(* IEC 61131-3 sources: LASAL/Class/SafetyCDIAS_Base (part 3) *)

	end_if;

END_FUNCTION

FUNCTION VIRTUAL SafetyCDIAS_Base::GetModuleID
	VAR_OUTPUT
		ud_ModuleID 	: UDINT;
	END_VAR

  // no module
  ud_ModuleID := 16#ff;

END_FUNCTION

FUNCTION VIRTUAL GLOBAL SafetyCDIAS_Base::Init
  VAR
		MyPara 	  : CmdStruct;
		MyResult	: results;
  END_VAR

//============================ Profiler start======================================================
#ifdef DM_Profiler
  InitTimeMeasurement(usMode := DMTIME_RT);
  InitTimeMeasurement(usMode := DMTIME_CY);
  InitTimeMeasurement(usMode := DMTIME_RTPOSTSCAN);
#endif
//============================ Profiler end========================================================

#ifdef DEACTIVATED_LSL
  IF Place.Read() = DEACTIVATED_LSL THEN
    State.uiIO_Flags                  := 0;
    State.uiIO_Flags.NoHW             := 1;
    State.uiIO_Flags.PhysicAccessOff  := 1;
    return;
  END_IF;
#endif

  case InitStep of
    0:
      // initialize HwBaseCDIAS
      if InitSafetyBase() then
        InitStep += 1;
      else
        //Remember flag that init failed, we must not try again otherwise the local var pSafetyManagerThis gets overwritten with nil if it already has been initialized
        InitStep := -1;
      end_if;

    1:
      // add update tasks in dependence on priority (prio 1 is added when us_FirstScan = 2, prio 2 @ us_FirstScan = 3...)
      if ( ( us_FirstScan - 1 ) = GetTaskPriority() ) then

        AddSafetyTask();

        InitStep += 1;

      end_if;

   2:
      // initialize safety module specific data (cpu, input, output) in last init and send OK to CPU

      if ((us_FirstScan = 10) & ((State.uiIO_Flags = 0 | DelayedStartup = 1))) then

        // log in to safety manager, if there is one
        if pSafetyManagerThis then
          MyPara.uiCmd    := CMD_SM_ADD_MODULE;
          MyPara.aPara[0] := ud_MyModuleID$DINT;
          MyPara.aPara[1] := THIS$DINT;
          pSafetyManagerThis^.NewInst(#MyPara, #MyResult);

          // check if quit error is avaialble
          MyPara.uiCmd    := CMD_SM_QUIT_ERROR_AVAILABLE;
          MyPara.aPara[0] := THIS$DINT;
          pSafetyManagerThis^.NewInst(#MyPara, #MyResult);

          // if the DLL has been found and the version shows that CDIAS safety is supported
          b_QuitErrorAvailable := (MyResult.aData[0]$DINT <> 0) & (MyResult.aData[4]$UDINT >= SAFETY_DLL_VERSION_CDIAS_QE);

          // give the manager more details about the module (if it didn't work at the first time and the safety number is valid)
          if (b_SafetyInfoOK = FALSE & ((DelayedStartup = 0) | ((DelayedStartup = 1 & SafetyNumber)))) then

            MyPara.uiCmd    := CMD_SM_ADD_MODULE_INFO;
            MyPara.aPara[0] := THIS$DINT;
            MyPara.aPara[1] := SafetyNumber$DINT;
            MyPara.aPara[2] := FW_Version$DINT;
            MyPara.aPara[3] := FPGA_Version$DINT;
            MyPara.aPara[4] := to_DINT(p_ObjectPath^$USINT) + 1; // size of path (length + 1 for the length information)
            MyPara.aPara[5] := p_ObjectPath$DINT;
            pSafetyManagerThis^.NewInst(#MyPara, #MyResult);
            b_SafetyInfoOK := MyResult.aData[0];
          end_if;
        else
          // if there is no manager, we don't have to wait in cywork until the initialisation is finished
          b_ManagerInitialisationFinished := TRUE;
          b_ManagerReadyForSDO            := TRUE;
        end_if;

        InitSafeModule();
      end_if;

    -1:
      //Error, nothing to do here, states are set before

  end_case;

  us_FirstScan += 1;

END_FUNCTION

FUNCTION VIRTUAL SafetyCDIAS_Base::GetTaskPriority
	VAR_OUTPUT
		us_TaskPriority 	: USINT;
	END_VAR

  // highest = default-priority (no change in update order)
  us_TaskPriority := 0;

END_FUNCTION

FUNCTION VIRTUAL SafetyCDIAS_Base::InitSafeModule
	VAR_OUTPUT
		sd_retval 	: DINT;
	END_VAR

  sd_retval := 0;

END_FUNCTION

FUNCTION VIRTUAL SafetyCDIAS_Base::StartDO
  VAR
  	i : DINT;
  END_VAR

  if b_PayloadSupport = FALSE then
    //set right address of do
    MasterConnect.SetNewDOAddressRd( p_data := pPDOReadData$^DINT, ud_address:= ( ui_MyPlace + OFFSET_SPDO_DATA ) );
  end_if;

  //start data object
  MasterConnect.ResetDO( p_data_object := p_HandlePDORead$^DINT, us_state := VARAN_DO_NO_RUN, ud_bytes := MaxLengthPDORead );

  // only for modules with outputs
  if Kennung <> CSDI16x_ID then
    if b_PayloadSupport = FALSE then
      //set right address of do
      MasterConnect.SetNewDOAddressWr( p_data := pPDOWriteData$^DINT, ud_address:= ( ui_MyPlace + OFFSET_SPDO_DATA ) );
    end_if;
    //start data object
    MasterConnect.ResetDO( p_data_object := p_HandlePDOWrite$^DINT, us_state := VARAN_DO_NO_RUN, ud_bytes := MaxLengthPDOWrite);

    if (AdditionalSPDOs > 0) then
      for i := 0 to (AdditionalSPDOs-1) do
        if b_PayloadSupport = FALSE then
          //set right address of do
          MasterConnect.SetNewDOAddressWr( p_data := aAdditionalPDOs[i].pPDOWriteData$^DINT, ud_address:= ( ui_MyPlace + OFFSET_SPDO_DATA ) );
        end_if;
        //start data object
        MasterConnect.ResetDO( p_data_object := aAdditionalPDOs[i].p_HandlePDOWrite$^DINT, us_state := VARAN_DO_NO_RUN, ud_bytes := MaxLengthPDOWrite);
      end_for;
    end_if;
  end_if;

  if b_PayloadSupport = FALSE then
    //set right address of do
    MasterConnect.SetNewDOAddressRd(p_data := p_us_Handle_TDO_Read$^DINT, ud_address := ui_MyPlace + OFFSET_STDO_DATA);

    //set right address of do
    MasterConnect.SetNewDOAddressWr(p_data := p_us_Handle_TDO_Write$^DINT, ud_address := ui_MyPlace + OFFSET_STDO_DATA);

    //set right address of do
    MasterConnect.SetNewDOAddressRd(p_data := p_ud_Handle_LED$^DINT, ud_address := ui_MyPlace + OFFSET_LED );
  end_if;

	//start data object
  MasterConnect.ResetDO( p_data_object := p_HandleTDORead$^DINT, us_state := VARAN_DO_NO_RUN, ud_bytes := STDO_LENGTH );

  //start data object
  MasterConnect.ResetDO( p_data_object := p_HandleTDOWrite$^DINT, us_state := VARAN_DO_NO_RUN, ud_bytes := STDO_LENGTH );

	//start data object
	MasterConnect.ResetDO( p_data_object := p_HandleLED$^DINT, us_state := VARAN_DO_CONT_RUN, ud_bytes := 15 );

  // only for modules with outputs
  if Kennung <> CSDI16x_ID then
    if b_PayloadSupport = FALSE then
      //set right address of do
      MasterConnect.SetNewDOAddressWr(p_data := p_ui_UnsafeOutWrite$^DINT, ud_address := ui_MyPlace + OFFSET_UNSAFE_VAR);
    end_if;
    //start data object
    MasterConnect.ResetDO( p_data_object := p_HandleUnsafeOutWrite$^DINT, us_state := VARAN_DO_NO_RUN, ud_bytes := UNSAFE_OUT_LENGTH );
  end_if;

  // fast unsafe variables (only if activated)
  if ActivateFastUnsafeIOs then
    if b_PayloadSupport = FALSE then
      //set right address of do
      MasterConnect.SetNewDOAddressRdWr(p_data:=p_us_Handle_FastUnsafeInputs$^DINT, ud_address_read:=ui_MyPlace + OFFSET_FAST_UNSAFE_IOS, ud_address_write:=ui_MyPlace + OFFSET_FAST_UNSAFE_IOS);
    end_if;
    //start data object
    MasterConnect.ResetDO( p_data_object := p_HandleFastUnsafeIOs$^DINT, us_state := VARAN_DO_CONT_RUN, ud_bytes := 1 );
  end_if;

  if b_PayloadSupport = FALSE then
    //set right address of do
    MasterConnect.SetNewDOAddressWr(p_data := p_us_Handle_TimeSyncHS_Write$^DINT, ud_address := ui_MyPlace + OFFSET_TIMESYNC_HANDSHAKE);
  end_if;
  //start data object
  MasterConnect.ResetDO( p_data_object := p_Handle_TimeSyncHS_Write$^DINT, us_state := VARAN_DO_NO_RUN, ud_bytes := 1 );

END_FUNCTION

FUNCTION VIRTUAL SafetyCDIAS_Base::StopDO
  VAR
  	i : DINT;
  END_VAR

  // stop data objects
	MasterConnect.ResetDO( p_data_object := p_HandlePDORead$^DINT, us_state := VARAN_DO_NO_RUN, ud_bytes := MaxLengthPDORead);

  // only for modules with outputs
  if Kennung <> CSDI16x_ID then

    MasterConnect.ResetDO( p_data_object := p_HandlePDOWrite$^DINT, us_state := VARAN_DO_NO_RUN, ud_bytes := MaxLengthPDOWrite);

    if (AdditionalSPDOs > 0) then
      for i := 0 to (AdditionalSPDOs-1) do
        if b_PayloadSupport = FALSE then
          //set right address of do
          MasterConnect.SetNewDOAddressWr( p_data := aAdditionalPDOs[i].pPDOWriteData$^DINT, ud_address:= ( ui_MyPlace + OFFSET_SPDO_DATA ) );
        end_if;
        //start data object
        MasterConnect.ResetDO( p_data_object := aAdditionalPDOs[i].p_HandlePDOWrite$^DINT, us_state := VARAN_DO_NO_RUN, ud_bytes := MaxLengthPDOWrite);
      end_for;
    end_if;
  end_if;

	MasterConnect.ResetDO( p_data_object := p_HandleTDORead$^DINT, us_state := VARAN_DO_NO_RUN, ud_bytes := STDO_LENGTH );
  b_DOIsRunningTDORead          := 0;

	MasterConnect.ResetDO( p_data_object := p_HandleTDOWrite$^DINT, us_state := VARAN_DO_NO_RUN, ud_bytes := STDO_LENGTH );
  b_DOIsRunningTDOWrite         := 0;

  MasterConnect.ResetDO( p_data_object := p_HandleLED$^DINT, us_state := VARAN_DO_NO_RUN, ud_bytes := 15 );

  MasterConnect.ResetDO( p_data_object := p_Handle_TimeSyncHS_Write$^DINT, us_state := VARAN_DO_NO_RUN, ud_bytes := 1 );
  b_DOIsRunning_TimeSyncHS      := 0;

  // only for modules with outputs
  if Kennung <> CSDI16x_ID then
    MasterConnect.ResetDO( p_data_object := p_HandleUnsafeOutWrite$^DINT, us_state := VARAN_DO_NO_RUN, ud_bytes := UNSAFE_OUT_LENGTH );
    b_DOIsRunningUnsafeOutWrite := 0;
  end_if;

END_FUNCTION

FUNCTION VIRTUAL SafetyCDIAS_Base::InitBuffers
	VAR_OUTPUT
		sd_retval 	: DINT;
	END_VAR

  sd_retval := -1;

  //allocate memory for outgoing SDO (one SDO possible)
  p_SDOOutputBuffer$^void := To_StdLib.Malloc(size := SDO_MAX_LENGTH);

  if ( p_SDOOutputBuffer = NIL ) then
    State.uiIO_Flags				          := 0;
		State.uiIO_Flags.PhysicAccessOff  := 1;
    ClassState := _MemAllocFailed;
    return;
  end_if;

  //allocate memory for incoming SDO list (number of SDO is dynamical)
  //following elements will be added dynamical

  //allocate list
  InputBufferAllocatedNo := SDO_BUFFER_ALLOC_BLOCK;
  p_SDOInputBuffer$^void := To_StdLib.Malloc(size := InputBufferAllocatedNo * SDO_MAX_LENGTH);

  if ( p_SDOInputBuffer = NIL ) then
    State.uiIO_Flags				          := 0;
		State.uiIO_Flags.PhysicAccessOff  := 1;
    ClassState := _MemAllocFailed;
    return;
  end_if;

  //all buffers initialized
  sd_retval := 0;

END_FUNCTION

FUNCTION VIRTUAL SafetyCDIAS_Base::GetSafetyNumber
	VAR_OUTPUT
		sd_retval 	: DINT;
	END_VAR
  VAR
  	TempPathInfo: PathInfoType;
		MyPara 	    : CmdStruct;
		MyResult	  : results;
  END_VAR

  sd_retval := SDOStdRequ ( us_Command      := SDO_COMMAND_GET_SAFENBR
                          , p_us_RespData   := ( #SafetyNumber )$^USINT
                          , us_RespLength   := sizeof(SafetyNumber)
                          );

  if ( sd_retval <> 0 ) then
    State.uiIO_Flags				          := 0;
		State.uiIO_Flags.PhysicAccessOff  := 1;

    LogError("@ZZZZ (SafetyCDIAS_Base::GetSafetyNumber) No Safety Number available!");
  elsif pConfigMem then
    // store safety number in config memory
    pConfigMem^$HDINT := SafetyNumber;
  end_if;

  sd_retval := SDOStdRequ ( us_Command      := SDO_COMMAND_GET_FW_VERSION
                          , p_us_RespData   := ( #FirmwareVersion )$^USINT
                          , us_RespLength   := sizeof(FirmwareVersionType)
                          );

  if ( sd_retval = 0 ) then
    FW_Version := FirmwareVersion.RevMinor OR (FirmwareVersion.RevMajor SHL 16);

    // Minor Versions starting with 9xxx mark Bootloader versions
    if (FirmwareVersion.RevMinor >= 9000) & (FirmwareVersion.RevMinor < 10000) then
      LogError("@ZZZZ (SafetyCDIAS_Base::GetSafetyNumber) Bootloader version of safety firmware detected! Download a firmware or contact Sigmatek Support!");
    end_if;

    // if we are connected over mover maybe the second try to read the fw version succeeds after the first failed
    if (sd_VaranType = 2) & (ClassState = _ReadFWVerFailed) then
      ClassState := _WaitForSynchronicity;
    end_if;
  else
    State.uiIO_Flags				          := 0;
    State.uiIO_Flags.PhysicAccessOff  := 1;
    ClassState := _ReadFWVerFailed;
    LogError("@ZZZZ (SafetyCDIAS_Base::GetSafetyNumber) No Firmware Version available!");
  end_if;

  InitPathInfo(#TempPathInfo);

  // add own safety number to routing table
  sd_retval := AddRoutingElement( ud_SafeNumber       := SafetyNumber
                                , ud_thisp            := this$UDINT
                                , pObject             := #TempPathInfo
                                );

  // give the manager more details about the module
  if pSafetyManagerThis then
    if ((SafetyNumber & DelayedStartup = 1) | DelayedStartup = 0) then
      MyPara.uiCmd    := CMD_SM_ADD_MODULE_INFO;
      MyPara.aPara[0] := THIS$DINT;
      MyPara.aPara[1] := SafetyNumber$DINT;
      MyPara.aPara[2] := FW_Version$DINT;
      MyPara.aPara[3] := FPGA_Version$DINT;
      MyPara.aPara[4] := to_DINT(p_ObjectPath^$USINT) + 1; // size of path (length + 1 for the length information)
      MyPara.aPara[5] := p_ObjectPath$DINT;
      pSafetyManagerThis^.NewInst(#MyPara, #MyResult);
      b_SafetyInfoOK := MyResult.aData[0];
    end_if;
  else
    // if there is no safety manager, it can only work if old modules are being used (new need the time sync token)

    // if the FPGA Version is lower than 1.4 or the minor firmware version is lower than 100 everything is fine
    if (FPGA_Version < 16#14) | (FW_Version$UINT < 100) then
      // new classes with old modules and without safety manager (hwcontrol) => no problem
    else
      // new classes with new modules and without safety manager (hwcontrol) => problem: noone there to pass on the time sync token
      LogError("@ZZZZ (SafetyCDIAS_Base::GetSafetyNumber) For new safety modules an object of HwControl is needed for time synchronisation!");
    end_if;
  end_if;

END_FUNCTION

FUNCTION SafetyCDIAS_Base::SafetyCDIAS_Base
	VAR_OUTPUT
		ret_code 	: ConfStates;
	END_VAR

#ifdef HWC_LogInit
  HWC_LogInit();
#endif

  //get interface for safety functions
  if ( OS_CILGET(INTERFACE_SAFETY, #pISafety)) then
    pISafety := NIL;

    LogError("@ZZZZ (SafetyCDIAS_Base::SafetyCDIAS_Base) No Safety Interface found!");

  end_if;

  // initialize it with FALSE, if there is anything on local CDIAS it will change to TRUE
  b_SafetyOnLocalCDIAS := FALSE;

  // initialize module count with 0
  ModuleSyncNo := 0;

  ret_code := C_OK;

END_FUNCTION

FUNCTION VIRTUAL GLOBAL SafetyCDIAS_Base::UpDateRT
	VAR_INPUT
		Handle 	      : UDINT;
	END_VAR
  VAR
    PDOLength     : USINT;
    p_ReceiveObj  : pVirtualBase;
    p_addressRd   : ^VaranDOSettingsRd;
    i             : DINT;
		MyPara 	      : CmdStruct;
		MyResult	    : results;
    bValidTDO     : BOOL;
  END_VAR

//============================ Profiler start======================================================
#ifdef  DM_Profiler
  StartTimeMeasurement(usMode := DMTIME_RT);
#endif
//============================ Profiler end========================================================

  // do tdo/pdo communication only, if module has been found and initialized correctly and if there are some LEDs on (else a FW-Update is running)
  if ( State.uiIO_Flags = 0 ) &
     (( ClassState = _SafetyClassOK ) | ( ClassState = _WaitForSynchronicity ) | ( ClassState = _ReinitConfig ) | ( ClassState = _ModFromCfgNotFound ) | ( ClassState = _UnknownCfgError ) | ( ClassState = _UnsafeVarNotFound )) then

    if StartRtDOs then
      if StartRtDOs = 2 then
        //start DOs
        StartDO();
      else
        if b_PayloadSupport = FALSE then
          //set right address of do
          MasterConnect.SetNewDOAddressRd( p_data := pPDOReadData$^DINT, ud_address:= ( ui_MyPlace + OFFSET_SPDO_DATA ) );
        end_if;

        //start data object
        MasterConnect.ResetDO( p_data_object := p_HandlePDORead$^DINT, us_state := VARAN_DO_NO_RUN, ud_bytes := MaxLengthPDORead );
      end_if;

      StartRtDOs := 0;
      return;
    end_if;

    // get I/O state, runstate, error
    UpDateNotStd(calloption:=CALL_OPTION_RT_PRESCAN);

    // wait until the safetymanager has initialized everything
    if b_ManagerInitialisationFinished = FALSE then
      return;
    end_if;

    // if any LED is active, then firmware update is not active and we can do our work
    if (VoltageOK | RunState | ServiceMode | Error) then
      // first check if there is a TDO to fetch
#ifdef SAFETY_OVER_DIAS
      if ( b_im ) then
        // Read Length of TDO
        TDOInfo := p_us_Handle_TDOReadLen^;

        // check msb (= new data) and length of frame
        if (TDOInfo AND 16#80) & ((TDOInfo AND 16#7F) = STDO_LENGTH) then

          //copy TDO word by word
          for i := 0 to (((TDOInfo AND 16#7F)/2)-1) by 1 do

            ( (#TDOFrame)$^UINT + ( i * 2 ) )^ := ( a_Handle_TDO_Read[i] )$^UINT^;

          end_for;

          // check length inside TDO Frame (must be 20)
          if TDOFrame.StdHeader.Len = 20 then

            // check who needs the TDO and give it the right addressee

            //search this-pointer of receiver with safety number
            p_ReceiveObj := ( GetRoutingPointerByNumber(ud_SafeNumber := TDOFrame.DstAdr))$pVirtualBase;

            if p_ReceiveObj <> NIL then
              MyPara.uiCmd := CMD_SM_WRITE_TDO_TO_MODULE;
              MyPara.aPara[0] := (#TDOFrame)$DINT;
              p_ReceiveObj^.NewInst(#MyPara, #MyResult);

  //                p_ReceiveObj^.WriteTDO2Module(#TDOFrame);
            end_if;
          else
            if bd_AlreadyLoggedMarker.TdoLenInvalid = FALSE then
              bd_LogOnceMarker.TdoLenInvalid := TRUE;
            end_if;
          end_if;
        end_if;
      else
#endif

        if NewHandShakeValue then

          p_us_Handle_TimeSyncHS_Write^ := p_us_Handle_TimeSyncHS_Read^ OR NewHandShakeValue;
          if b_VaranAvailable then

            if b_PayloadSupport then
              if sd_VaranType = 2 then
                p_Handle_TimeSyncHS_WriteEnable^ := VARAN_MOVER_DO_CONT_RUN;
                TimeSyncHSSingleRunActive := 2;
              else
                b_DOIsRunning_TimeSyncHS.StartRequest := true;
              end_if;
            else
              if sd_VaranType = 2 then
                (p_Handle_TimeSyncHS_Write$^USINT )^ := VARAN_MOVER_DO_CONT_RUN;
                TimeSyncHSSingleRunActive := 2;
              else
                MasterConnect.ResetDO( p_data_object := p_Handle_TimeSyncHS_Write$^DINT, us_state := VARAN_DO_SINGLE_RUN, ud_bytes := 1 );
              end_if;
            end_if;

          end_if;

          // if the time synchonisation is active we send 2 different bits in 2 successive cycles, so the µC can detect the cycle time
          if NewHandShakeValue = 2#011 then
            NewHandShakeValue := 2#111;
            if sd_VaranType = 1 then
              // start DO at this point to ensure 1 cycle delay, from request to response
              if b_PayloadSupport then
                EnableDO(ud_DOHandle := p_HandleTDORead$UDINT);
                b_DOIsRunningTDORead.ContRun := true;
              else
                p_HandleTDORead^.ucCtrlStat := VARAN_DO_CONT_RUN;
              end_if;

            end_if;
            TimeSyncDOActive.OwnSyncActive := 1;
          else
            NewHandShakeValue := 0;
          end_if;
        elsif b_TimeSyncActive then
          // on input or output module we wait until the time synchronisation is finished
          if ((p_us_Handle_TimeSyncHS_Read^ AND 2#110) = 0) & (TimeSyncHSSingleRunActive = 0) then
            b_TimeSyncActive := FALSE;
            TimeSyncDOActive.OwnSyncActive := 0;

            // if we have no mover and no external request is pending => stop the read DO
            if (sd_VaranType = 1) & (TimeSyncDOActive$DINT = 0) then

              if b_PayloadSupport then

                if b_DOIsRunningTDORead = 0 then
                  if bd_AlreadyLoggedMarker.TdoLenInvalid = FALSE then
                    bd_LogOnceMarker.TdoLenInvalid := TRUE;
                  end_if;
                end_if;
                DisableDO(ud_DOHandle := p_HandleTDORead$UDINT);
                b_DOIsRunningTDORead := 0;

              else

                if p_HandleTDORead^.ucCtrlStat AND 0x03 = VARAN_DO_NO_RUN then
                  if bd_AlreadyLoggedMarker.TdoLenInvalid = FALSE then
                    bd_LogOnceMarker.TdoLenInvalid := TRUE;
                  end_if;
                end_if;
                p_HandleTDORead^.ucCtrlStat := VARAN_DO_NO_RUN;

              end_if;

            end_if;
            MyPara.uiCmd := CMD_SM_TIME_SYNC_FINISHED;
            pSafetyManagerThis^.NewInst(#MyPara, #MyResult); // thispointer doesn't have to be checked here; NewHandShakeValue gets set via SafetyManager
          end_if;
        end_if;

        // Read Length of TDO
        TDOInfo := p_us_Handle_TDO_Read_Length^;

        // check msb (= new data) and length of frame
        bValidTDO := (TDOInfo AND 16#80) & ((TDOInfo AND 16#7F) = STDO_LENGTH);

        if b_VaranAvailable then

          if (sd_VaranType = 1) then // ----------------------------------------------------------------------

            if b_NewSyncMode then
              if bValidTDO then
                if b_PayloadSupport then

                // check if data-DO is running already
                  if b_DOIsRunningTDORead.ContRun then
                    TDOTransStarted := TRUE;
                  else
                    // we didn´t expect this, so read out and ignore (maybe its an old frame)
                    b_DOIsRunningTDORead.StartRequest := true;
                    bValidTDO := FALSE;
                  end_if;

                else

                    // check if data-DO is running already
                  if (p_HandleTDORead^.ucCtrlStat AND 16#03) = VARAN_DO_CONT_RUN then
                    TDOTransStarted := TRUE;
                  else
                    // we didn´t expect this, so read out and ignore (maybe its an old frame)
                    p_HandleTDORead^.ucCtrlStat := VARAN_DO_SINGLE_RUN;
                    bValidTDO := FALSE;
                  end_if;

                end_if;
              end_if;
            end_if;

            // if we got the TDO Data, copy them
            if TDOTransStarted then

              //copy whole TDO
              To_StdLib.MemCpy(dest := #TDOFrame, source := p_us_Handle_TDO_Read, size := sizeof(TDOType));

#ifdef SAFETY_PROTOCOL_ANALYZER_ACTIVATED
  RecordFrame((#TDOFrame)$^DINT, 0);
#endif

              // check length inside TDO Frame (must be 20)
              if TDOFrame.StdHeader.Len = (STDO_LENGTH - sizeof(TDOType.StdHeader.CRC)) then
                TDOTransStarted := FALSE;

                // if our own timesynchronisation is not running => stop the read DO
                if b_NewSyncMode & (TimeSyncDOActive$DINT = 0) then
                  if b_PayloadSupport then
                    DisableDO(ud_DOHandle := p_HandleTDORead$UDINT);  // we got data, so stop DO
                    b_DOIsRunningTDORead := 0;
                  else
                    p_HandleTDORead^.ucCtrlStat := VARAN_DO_NO_RUN; // we got data, so stop DO
                  end_if;
                end_if;
                // check who needs the TDO and give it the right addressee

                //search this-pointer of receiver with safety number
                p_ReceiveObj := ( GetRoutingPointerByNumber(ud_SafeNumber := TDOFrame.DstAdr))$pVirtualBase;

                if p_ReceiveObj <> NIL then
#ifdef DO_DEBUG
                  DOCheck(pFrame:=(#TDOFrame)$^SDOStdHeader, pCheckStruct:=#TDORead);
#endif

                  MyPara.uiCmd    := CMD_SM_WRITE_TDO_TO_MODULE;
                  MyPara.aPara[0] := (#TDOFrame)$DINT;
                  p_ReceiveObj^.NewInst(#MyPara, #MyResult);

  //                p_ReceiveObj^.WriteTDO2Module(#TDOFrame);
                elsif pSafetyManagerThis then
#ifdef DO_DEBUG
                  DOCheck(pFrame:=(#TDOFrame)$^SDOStdHeader, pCheckStruct:=#TDORead);
#endif

                  //passing the TDO to another domain
                  MyPara.uiCmd    := CMD_SM_TDO_TO_MANAGER;
                  MyPara.aPara[0] := STDO_LENGTH;
                  MyPara.aPara[1] := (#TDOFrame)$DINT;
                  pSafetyManagerThis^.NewInst(#MyPara, #MyResult);
                end_if;
              elsif TDOFrame.StdHeader.Len > 0 then
                if bd_AlreadyLoggedMarker.TdoLenInvalid = FALSE then
                  bd_LogOnceMarker.TdoLenInvalid := TRUE;
                end_if;
              end_if;
            end_if;

            if (b_NewSyncMode = FALSE) & (TDOInfo AND 16#80) then
              if ((TDOInfo AND 16#7F) = STDO_LENGTH) then

                // if so, start DO and remember to use info next time
                if b_PayloadSupport then
                  b_DOIsRunningTDORead.StartRequest := true;
                else
                  p_HandleTDORead^.ucCtrlStat := VARAN_DO_SINGLE_RUN;
                end_if;

                if ((TDOFrame.StdHeader.Typ AND SSDO_MASK_RESPONSE) = 0) & (udTDORdCnt < 2) then
                  udTDORdCnt += 1;
                else
                  TDOTransStarted := TRUE;
                end_if;
              end_if;
            end_if;
          else  // Mover active ----------------------------------------------------------------------
            if TimeSyncHSSingleRunActive then
              TimeSyncHSSingleRunActive -= 1;
              if TimeSyncHSSingleRunActive = 0 then
                if b_PayloadSupport then
                  p_Handle_TimeSyncHS_WriteEnable^      := VARAN_DO_NO_RUN;
                else
                  (p_Handle_TimeSyncHS_Write$^USINT )^  := VARAN_DO_NO_RUN;
                end_if;
              end_if;
            end_if;

            if bValidTDO then

              //copy whole TDO
              To_StdLib.MemCpy(dest := #TDOFrame, source := p_us_Handle_TDO_Read, size := sizeof(TDOType));

#ifdef SAFETY_PROTOCOL_ANALYZER_ACTIVATED
RecordFrame((#TDOFrame)$^DINT, 0);
#endif

              // check length inside TDO Frame (must be 20)
              if TDOFrame.StdHeader.Len = (STDO_LENGTH - sizeof(TDOType.StdHeader.CRC)) then

                // check who needs the TDO and give it the right addressee

                //search this-pointer of receiver with safety number
                p_ReceiveObj := ( GetRoutingPointerByNumber(ud_SafeNumber := TDOFrame.DstAdr))$pVirtualBase;

                if p_ReceiveObj <> NIL then
#ifdef DO_DEBUG
                  DOCheck(pFrame:=(#TDOFrame)$^SDOStdHeader, pCheckStruct:=#TDORead);
#endif

                  MyPara.uiCmd    := CMD_SM_WRITE_TDO_TO_MODULE;
                  MyPara.aPara[0] := (#TDOFrame)$DINT;
                  p_ReceiveObj^.NewInst(#MyPara, #MyResult);

      //                p_ReceiveObj^.WriteTDO2Module(#TDOFrame);
                elsif pSafetyManagerThis then
#ifdef DO_DEBUG
                  DOCheck(pFrame:=(#TDOFrame)$^SDOStdHeader, pCheckStruct:=#TDORead);
#endif

                  //passing the TDO to another domain
                  MyPara.uiCmd    := CMD_SM_TDO_TO_MANAGER;
                  MyPara.aPara[0] := STDO_LENGTH;
                  MyPara.aPara[1] := (#TDOFrame)$DINT;
                  pSafetyManagerThis^.NewInst(#MyPara, #MyResult);
                end_if;
              elsif TDOFrame.StdHeader.Len > 0 then
                if bd_AlreadyLoggedMarker.TdoLenInvalid = FALSE then
                  bd_LogOnceMarker.TdoLenInvalid := TRUE;
                end_if;
              elsif TDOFrame.StdHeader.Len = 0 then
                if bd_AlreadyLoggedMarker.TdoLen0 = FALSE then
                  bd_LogOnceMarker.TdoLen0 := TRUE;
                end_if;
              end_if;
            end_if;
          end_if; // --------------------------------------------------------------------------------------
        else  // if b_VaranAvailable then
          if bValidTDO then

            //copy whole TDO
            To_StdLib.MemCpy(dest := #TDOFrame, source := p_us_Handle_TDO_Read, size := sizeof(TDOType));

#ifdef DO_DEBUG
            DOCheck(pFrame:=(#TDOFrame)$^SDOStdHeader, pCheckStruct:=#TDORead);
#endif

#ifdef SAFETY_PROTOCOL_ANALYZER_ACTIVATED
  RecordFrame((#TDOFrame)$^DINT, 0);
#endif

            // check length inside TDO Frame (must be 20)
            if TDOFrame.StdHeader.Len = (STDO_LENGTH - sizeof(TDOType.StdHeader.CRC)) then

              // check who needs the TDO and give it the right addressee

              //search this-pointer of receiver with safety number
              p_ReceiveObj := ( GetRoutingPointerByNumber(ud_SafeNumber := TDOFrame.DstAdr))$pVirtualBase;

              if p_ReceiveObj <> NIL then
                if ((TDOFrame.StdHeader.Typ AND SSDO_MASK_RESPONSE) = 0) & (udTDORdCnt < 2) then
                  udTDORdCnt += 1;
                else
#ifdef DO_DEBUG
                  DOCheck(pFrame:=(#TDOFrame)$^SDOStdHeader, pCheckStruct:=#TDORead);
#endif

                  MyPara.uiCmd    := CMD_SM_WRITE_TDO_TO_MODULE;
                  MyPara.aPara[0] := (#TDOFrame)$DINT;
                  p_ReceiveObj^.NewInst(#MyPara, #MyResult);

      //                p_ReceiveObj^.WriteTDO2Module(#TDOFrame);
                end_if;
              elsif pSafetyManagerThis then
#ifdef DO_DEBUG
                DOCheck(pFrame:=(#TDOFrame)$^SDOStdHeader, pCheckStruct:=#TDORead);
#endif

                //passing the TDO to another domain
                MyPara.uiCmd    := CMD_SM_TDO_TO_MANAGER;
                MyPara.aPara[0] := STDO_LENGTH;
                MyPara.aPara[1] := (#TDOFrame)$DINT;
                pSafetyManagerThis^.NewInst(#MyPara, #MyResult);
              end_if;
            else
              if bd_AlreadyLoggedMarker.TdoLenInvalid = FALSE then
                bd_LogOnceMarker.TdoLenInvalid := TRUE;
              end_if;
            end_if;
          end_if;
        end_if;

        if bValidTDO then
          // if it's a response, reset the flag
          if TDOFrame.StdHeader.Typ AND 16#80 then
            TimeSyncDOActive.Wait4ResponseNo -= 1;
          end_if;
        end_if;

#ifdef SAFETY_OVER_DIAS
      end_if;
#endif

      // if we are in run state
      if RunState then

        // we have to start the DOs here because it's the right task for this
        if b_StartDOs then
          b_StartDOs := FALSE;
          if sd_VaranType = 1 then
            if b_PayloadSupport = FALSE then
              //set right address of do
              MasterConnect.SetNewDOAddressWr( p_data := pPDOWriteData$^DINT, ud_address:= ( ui_MyPlace + OFFSET_SPDO_DATA ) );
            end_if;

            MasterConnect.ResetDO( p_data_object := p_HandlePDOWrite$^DINT, us_state := VARAN_DO_CONT_RUN, ud_bytes := MaxLengthPDOWrite);

            if AdditionalSPDOs & (ui_cnt_PDOInputBuffer > 1) then
              if AdditionalSPDOs > (ui_cnt_PDOInputBuffer-1) then
                AdditionalSPDOs := ui_cnt_PDOInputBuffer-1;
              end_if;

              for i := 0 to (AdditionalSPDOs-1) do
                if b_PayloadSupport = FALSE then
                  //set right address of do
                  MasterConnect.SetNewDOAddressWr( p_data := aAdditionalPDOs[i].pPDOWriteData$^DINT, ud_address:= ( ui_MyPlace + OFFSET_SPDO_DATA ) );
                end_if;

                MasterConnect.ResetDO( p_data_object := aAdditionalPDOs[i].p_HandlePDOWrite$^DINT, us_state := VARAN_DO_CONT_RUN, ud_bytes := MaxLengthPDOWrite);
              end_for;
            end_if;
          else

            if b_PayloadSupport then
              p_HandlePDOWriteEnable^     := VARAN_MOVER_DO_CONT_RUN; // = VARAN_DO_SINGLE_RUN
            else
              (p_HandlePDOWrite$^USINT )^ := VARAN_MOVER_DO_CONT_RUN; // is continous at the mover
            end_if;

            if AdditionalSPDOs & (ui_cnt_PDOInputBuffer > 1) then
              if AdditionalSPDOs > (ui_cnt_PDOInputBuffer-1) then
                AdditionalSPDOs := ui_cnt_PDOInputBuffer-1;
              end_if;

              for i := 0 to (AdditionalSPDOs-1) do
                if b_PayloadSupport then
                  aAdditionalPDOs[i].p_HandlePDOWriteEnable^    := VARAN_MOVER_DO_CONT_RUN; // = VARAN_DO_SINGLE_RUN
                else
                  (aAdditionalPDOs[i].p_HandlePDOWrite$^USINT )^:= VARAN_MOVER_DO_CONT_RUN; // is continous at the mover
                end_if;
              end_for;
            end_if;
          end_if;
        end_if;

        if b_MoveCommandOutputActive <> _Active then
          if PDOSingleRunActive then
            PDOSingleRunActive -= 1;
            if PDOSingleRunActive = 0 then

              if b_PayloadSupport then  // ---------------------------------

                if (sd_VaranType = 1) then  // Payload Without Mover +++++++
                  DisableDO(ud_DOHandle := p_HandlePDOWrite$UDINT);

                  if AdditionalSPDOs then
                    for i := 0 to (AdditionalSPDOs-1) do
                      DisableDO(ud_DOHandle := aAdditionalPDOs[i].p_HandlePDOWrite$UDINT );
                    end_for;
                  end_if;

                else  // Payload With Mover ++++++++++++++++++++++++++++++++
                  p_HandlePDOWriteEnable^ := VARAN_DO_NO_RUN;

                  if AdditionalSPDOs then
                    for i := 0 to (AdditionalSPDOs-1) do
                      (aAdditionalPDOs[i].p_HandlePDOWriteEnable)^ := VARAN_DO_NO_RUN;
                    end_for;
                  end_if;
                end_if; // +++++++++++++++++++++++++++++++++++++++++++++++++

              else  // No Payload Wih Mover --------------------------------
                (p_HandlePDOWrite$^USINT )^ := VARAN_DO_NO_RUN;

                if AdditionalSPDOs then
                  for i := 0 to (AdditionalSPDOs-1) do
                    (aAdditionalPDOs[i].p_HandlePDOWrite$^USINT )^ := VARAN_DO_NO_RUN;
                  end_for;
                end_if;
              end_if; // ---------------------------------------------------

            end_if;
          end_if;

          //read PDO from hardware, only if PDO is needed by other moduls
          if ( PDOOutputIsUsed ) then
#ifdef SAFETY_OVER_DIAS
            if ( b_im ) then

              PDOLength := p_us_Handle_PDOReadLen^;

              // only if length is bigger than minimum and smaller than maximum
              if ( PDOLength > PDOType.Length ) & ( PDOLength <= SPDO_MAX_LENGTH) then
                //copy PDO word by word
                for i := 0 to ((PDOLength/2)-1) by 1 do

                  ( p_PDOOutputBuffer$^UINT + ( i * 2 ) )^ := ( a_Handle_PDO_Read[i] )$^UINT^;

                end_for;
              end_if;
            else
#endif

              PDOLength := pPDOReadLengthData^;

              if b_VaranAvailable & (sd_VaranType = 1) then

                // if "pdo length" matches the length of Varan-PDO data object
                if PDOLength = PDOReadLen then
                  // only if length is bigger than minimum and smaller than maximum
                  if ( PDOLength > PDOType.Length ) & ( PDOLength <= SPDO_MAX_LENGTH) then
                    //copy whole PDO
                    To_StdLib.MemCpy(dest := #PDOOutputBuffer, source := pPDOReadData, size := PDOLength);

#ifdef DO_DEBUG
                    DOCheck(pFrame:=(#PDOOutputBuffer)$^SDOStdHeader, pCheckStruct:=#PDORead);
#endif

#ifdef SAFETY_PROTOCOL_ANALYZER_ACTIVATED
//if ClassState = _SafetyClassOK then
  RecordFrame((#PDOOutputBuffer)$^DINT, 0);
//end_if;
#endif

                  end_if;
                else

                  if b_PayloadSupport then
                  // correct size of data object to PDOLength
                    ChangeDOLengthOffset( ud_DOHandle     := p_HandlePDORead$UDINT
                                        , ud_length_read  := PDOLength
                                        );
                    PDOReadLen              := PDOLength;
                    EnableDO(ud_DOHandle    := p_HandlePDORead$UDINT);
                  else
                    // correct size of data object to PDOLength
                    p_addressRd             := pPDOReadData - sizeof(VaranDOSettingsRd);
                    p_addressRd^.us_ByteCnt := PDOLength;
                    p_HandlePDORead^.usLengthofExpAnswer := sizeof(VaranDOSettingsRd.us_Command) + to_uint(PDOLength);

                    PDOReadLen := PDOLength;

                    MasterConnect.ResetDO( p_data_object := p_HandlePDORead$^DINT, us_state := VARAN_DO_CONT_RUN, ud_bytes := PDOLength );
                  end_if;

                end_if;
              else
                // only if length is bigger than minimum and smaller than maximum
                if ( PDOLength > PDOType.Length ) & ( PDOLength <= SPDO_MAX_LENGTH) then
                  //copy whole PDO
                  To_StdLib.MemCpy(dest := #PDOOutputBuffer, source := pPDOReadData, size := PDOLength);

#ifdef DO_DEBUG
                  DOCheck(pFrame:=(#PDOOutputBuffer)$^SDOStdHeader, pCheckStruct:=#PDORead);
#endif

#ifdef SAFETY_PROTOCOL_ANALYZER_ACTIVATED
//if ClassState = _SafetyClassOK then
  RecordFrame((#PDOOutputBuffer)$^DINT, 0);
//end_if;
#endif

                end_if;
              end_if;
#ifdef SAFETY_OVER_DIAS
            end_if;
#endif
          end_if;
        else
          PDOLength := pPDOReadLengthData^;

          // if "pdo length" doesn't match the length of Varan-PDO data object
          if (PDOLength <> PDOReadLen) & (sd_VaranType = 1) & ( PDOLength > PDOType.Length ) & ( PDOLength <= SPDO_MAX_LENGTH) then

            if b_PayloadSupport then
            // correct size of data object to PDOLength
              ChangeDOLengthOffset( ud_DOHandle     := p_HandlePDORead$UDINT
                                  , ud_length_read  := PDOLength
                                  );

              PDOReadLen := PDOLength;

              EnableDO(ud_DOHandle := p_HandlePDORead$UDINT);
            else
              // correct size of data object to PDOLength
              p_addressRd := pPDOReadData - sizeof(VaranDOSettingsRd);
              p_addressRd^.us_ByteCnt := PDOLength;
              p_HandlePDORead^.usLengthofExpAnswer := sizeof(VaranDOSettingsRd.us_Command) + to_uint(PDOLength);

              PDOReadLen := PDOLength;

              if b_PayloadSupport = FALSE then
                //set right address of do
                MasterConnect.SetNewDOAddressRd( p_data := pPDOReadData$^DINT, ud_address:= ( ui_MyPlace + OFFSET_SPDO_DATA ) );
              end_if;

              MasterConnect.ResetDO( p_data_object := p_HandlePDORead$^DINT, us_state := VARAN_DO_CONT_RUN, ud_bytes := PDOLength );
            end_if;

          end_if;

#ifdef DO_DEBUG
          DOCheck(pFrame:=pPDOReadData$^SDOStdHeader, pCheckStruct:=#PDORead);
#endif
        end_if;
      end_if;
    end_if;
  end_if;

  if b_PayloadSupport & (sd_VaranType = 1) then

    // s_DO_AcyRd xxxxxxxxxxxxxxxxxxxxxxxxxxxxxxxxxxxxxxxxxxxxxxxxxxxxxxxxxxxxxxxxxxxxxxxxxxxxxxxxxxxxxxxxxxxxxxxx
    case b_DOIsRunning_TimeSyncHS of

      SR_STATE_ENABLE_ME :  // DO is not running and start request is set ----------------------------------------
        EnableDO(ud_DOHandle := p_Handle_TimeSyncHS_Write$UDINT);
        b_DOIsRunning_TimeSyncHS := SR_STATE_DISABLE_ME;

      SR_STATE_DISABLE_ME : // DO is running and start request is not set ----------------------------------------
        DisableDO(ud_DOHandle:= p_Handle_TimeSyncHS_Write$UDINT);
        b_DOIsRunning_TimeSyncHS := SR_STATE_NOTHING;

      SR_STATE_LEAVE_ME_ENABLED : // DO is running and another start request is set ------------------------------
        b_DOIsRunning_TimeSyncHS := SR_STATE_DISABLE_ME;

    end_case;

  end_if;

#ifndef CALL_OPTION_RT_POSTSCAN
  UpDateRTPostScan(Handle);
#endif

//============================ Profiler start======================================================
#ifdef  DM_Profiler
  StopTimeMeasurement(usMode := DMTIME_RT);
#endif
//============================ Profiler end========================================================

END_FUNCTION

#pragma warning(disable:0073);
FUNCTION VIRTUAL SafetyCDIAS_Base::UpDateNotStd
	VAR_INPUT
		calloption 	: UDINT;
	END_VAR

END_FUNCTION
#pragma warning(default:0073);

FUNCTION VIRTUAL SafetyCDIAS_Base::ReadSDOConfig
	VAR_INPUT
		p_SDORequestBuffer 	          : ^SDORequReadConfig;
		p_SDOResponseBuffer 	        : ^SDORespReadConfig;
		pModule 	                    : ^PathInfoType;
		pListHeader 	                : ^PathInfoType;
	END_VAR
	VAR_OUTPUT
		sd_retval 	                  : DINT;
	END_VAR
  VAR
    ud_Address                    : UDINT;
    ud_ListLength_Address         : UDINT;
    ud_ListLength                 : UDINT;
    ud_TmpCnt                     : UDINT;
    i                             : UDINT;
    ud_ModulePathLen_Max          : UDINT;
    ud_ModulePathCompLen_Max      : UDINT;
    ud_ListHeaderPathLen_Max      : UDINT;
    ud_ListHeaderPathCompLen_Max  : UDINT;
    us_DataLength_Max             : USINT;
    ud_ListBaseAddress            : UDINT;
    ud_ListAddressMax             : UDINT;
    ud_CntUnsafeOutputs           : UDINT;
    ud_CntUnsafeInputs            : UDINT;
    ud_ActAddress                 : UDINT;  // actual offset in application memory (where to find the values in run mode)
    ud_UnsafeBDINT_Offset         : UDINT;  // actual offset in application memory (where to find the unsafe variables in run mode)
    ud_ActBlockType               : UDINT;
    ud_TmpAddress                 : UDINT;
    ud_TmpStrLen                  : UDINT;
    p_TmpBlockedData              : ^void;
    ud_ActStrLen                  : UDINT;
    us_BlockedTransferLength      : USINT;
    BoolOuts                      : UDINT;
    DintOuts                      : UDINT;
    TempModuleConfig              : t_ModuleCfg;
    pChar                         : ^CHAR;
    TempPath                      : ARRAY [0..99] OF USINT;
    PathOfThisCPU                 : ARRAY [0..99] OF USINT;
    GotOwnPath                    : BOOL;
    TempPdoConfig                 : t_PdoCfg;
    pBitMasks                     : ^BDINT;
    ActBitMask                    : BDINT;
    ud_skipLength                 : UDINT; //++pr
    b_CfgTypeV2                   : BOOL; // FALSE means there is no support of new time synchronisation/new general purpose register
    TmpCRC                        : HDINT;
    ud_ContainerBlockType         : UDINT;
    b_CfgTypeV3                   : BOOL;
    ud_ConfigLength               : UDINT;
    hd_DynParaVersion             : UDINT;
  END_VAR

  // Initialize the variables with invalid if we are located on VARAN. If any module to communicate with is not located on VARAN, it will change to inactive. (ConfigSafetyInput/Output)
  if b_VaranAvailable then
    b_MoveCommandInputActive    := _Invalid;
    b_MoveCommandOutputActive   := _Invalid;
  else
    // if no VARAN, we can't move the PDOs
    b_MoveCommandInputActive    := _Inactive;
    b_MoveCommandOutputActive   := _Inactive;
  end_if;

  //minimum length of path: 2 bytes length, 1 byte domain info, 1 byte bus type and 1 byte port
  ud_ModulePathLen_Max          := 5;
  ud_ModulePathCompLen_Max      := 5;
  ud_ListHeaderPathLen_Max      := 5;
  ud_ListHeaderPathCompLen_Max  := 5;

  NewConfigType                 := ConfigState_NotInitialized;

  //initialize header-data for request

  //calculate length without crc
  p_SDORequestBuffer^.StdHeader.Len := sizeof(SDORequReadConfig) - sizeof(SDOHeader.StdHeader.CRC);

  //type
  p_SDORequestBuffer^.StdHeader.Typ := SDO_STD;

  //command for reading config data
  p_SDORequestBuffer^.StdHeader.Cmd := SDO_COMMAND_READ;

  //read crc of whole config data

  //send request and receive data
  sd_retval := SDOReadCfgRequ ( p_SDORequestBuffer  := p_SDORequestBuffer
                              , p_SDOResponseBuffer := p_SDOResponseBuffer
                              , ud_Address          := SDO_ADDRESS_CONFIG_DATA + SDO_OFFSET_CONFIG_CRC_ALL
                              , us_Length           := 4
                              );

  //no response
  if ( sd_retval <> 0 ) then
    LogError("@ZZZZ (SafetyCDIAS_Base::ReadSDOConfig) Config Read Error: Error reading CRC of config data");
    return;
  end_if;

  // save crc and remember the time
  ud_ConfigCRC          := p_SDOResponseBuffer^.ud_Data;
  //Show CRC on Server
  DesignerPrjConfigCRC  := ud_ConfigCRC;
  ud_LastCrcCheck       := ops.tAbsolute;
  b_CheckCRC            := TRUE;

  //read length of whole config data

  //send request and receive data
  sd_retval := SDOReadCfgRequ ( p_SDORequestBuffer  := p_SDORequestBuffer
                              , p_SDOResponseBuffer := p_SDOResponseBuffer
                              , ud_Address          := SDO_ADDRESS_CONFIG_DATA + SDO_OFFSET_CONFIG_LEN_ALL
                              , us_Length           := 4
                              );

  //no response
  if ( sd_retval <> 0 ) then
    LogError("@ZZZZ (SafetyCDIAS_Base::ReadSDOConfig) Config Read Error: Error reading length of config data");
    return;
  end_if;

  //no config data available
  if ( p_SDOResponseBuffer^.ud_Data = 16#FFFF_FFFF ) then
    LogError("@ZZZZ (SafetyCDIAS_Base::ReadSDOConfig) Config Read Error: No config data available.");
    return;
  end_if;

  ud_ConfigLength := p_SDOResponseBuffer^.ud_Data;

  // get BlockType
  //send request and receive data
  sd_retval := SDOReadCfgRequ ( p_SDORequestBuffer  := p_SDORequestBuffer
                              , p_SDOResponseBuffer := p_SDOResponseBuffer
                              , ud_Address          := SDO_ADDRESS_CONFIG_DATA + SDO_OFFSET_CONFIG_BLOCKTYPE
                              , us_Length           := 4
                              );
  //no response, error
  if ( sd_retval <> 0 ) then
    LogError("@ZZZZ (SafetyCDIAS_Base::ReadSDOConfig) Config Read Error: Error getting the block type of the header");
    return;
  end_if;

  ud_ContainerBlockType := p_SDOResponseBuffer^.ud_Data;

  // check if it's a new version of the configuration
  if (ud_ContainerBlockType = BLKTYPE_CFG_CONTAINER_V3)       |
     (ud_ContainerBlockType = BLKTYPE_CFG_CONTAINER_V3_SLAVE)     |
     (ud_ContainerBlockType = BLKTYPE_CFG_CONTAINER_V3_SLAVE_OPTIONAL) then

    //read dynamic header length (how many data are attached to the header)

    //send request and receive data
    sd_retval := SDOReadCfgRequ ( p_SDORequestBuffer  := p_SDORequestBuffer
                                , p_SDOResponseBuffer := p_SDOResponseBuffer
                                , ud_Address          := SDO_ADDRESS_CONFIG_DATA + SDO_OFFSET_CONFIG_LEN_HEAD
                                , us_Length           := 4
                                );

    //no response
    if ( sd_retval <> 0 ) then
      LogError("@ZZZZ (SafetyCDIAS_Base::ReadSDOConfig) Config Read Error: Error reading length of dynamic header data");
      return;
    end_if;

    // plausibility check for data length
    if p_SDOResponseBuffer^.ud_Data > 1000 then
      sd_retval := -1;
      LogError("@ZZZZ (SafetyCDIAS_Base::ReadSDOConfig) Config Read Error: Invalid length of dynamic header data");
      return;
    end_if;

    // the length info contains: size of length info + size of time info + size of additional data

    //start address of first list: address of dynamic length + length according to length info
    ud_ListBaseAddress := SDO_ADDRESS_CONFIG_DATA + SDO_OFFSET_CONFIG_LEN_HEAD + p_SDOResponseBuffer^.ud_Data;

    // if we got at least 4 byte additional header data, it's the version of the dynamic parameters => read it
    if p_SDOResponseBuffer^.ud_Data >= 12 then
      //send request and receive data
      sd_retval := SDOReadCfgRequ ( p_SDORequestBuffer  := p_SDORequestBuffer
                                  , p_SDOResponseBuffer := p_SDOResponseBuffer
                                  , ud_Address          := SDO_ADDRESS_CONFIG_DATA + SDO_OFFSET_CONFIG_LEN_HEAD + 8
                                  , us_Length           := 4
                                  );

      //no response
      if ( sd_retval <> 0 ) then
        LogError("@ZZZZ (SafetyCDIAS_Base::ReadSDOConfig) Config Read Error: Error reading length of dynamic header data");
        return;
      end_if;

      hd_DynParaVersion := p_SDOResponseBuffer^.ud_Data;
    else
      LogError("@ZZZZ (SafetyCDIAS_Base::ReadSDOConfig) Config Read Error: Data structure error in config! No bytes for the dynamic parameter version (according to length info)!");
      return;
    end_if;
  else
    // old version => no dynamic header, the first list starts where the dynamic header length would be

    //start address of first list: address of time info + size of time info
    ud_ListBaseAddress := SDO_ADDRESS_CONFIG_DATA + SDO_OFFSET_CONFIG_LEN_HEAD + sizeof(UDINT);
  end_if;

  GotOwnPath := FALSE;

  //highest address for config data
  ud_ListAddressMax := SDO_ADDRESS_CONFIG_DATA + SDO_OFFSET_CONFIG_LEN_ALL + ud_ConfigLength;

  //max. length of data to read with one request
  us_DataLength_Max := SDO_MAX_LENGTH - sizeof(SDORespReadConfig) + sizeof(SDORespReadConfig.ud_Data);

  while ( ud_ListBaseAddress < ud_ListAddressMax ) do

    //first read length of path in list-header

    //read path in list-header
    sd_retval := ReadModulePath ( p_SDORequestBuffer          := p_SDORequestBuffer
                                , p_SDOResponseBuffer         := p_SDOResponseBuffer
                                , p_ud_Address                := #ud_ListBaseAddress
                                , pModule                     := pListHeader
                                , p_ud_ModulePathLen_Max      := #ud_ListHeaderPathLen_Max
                                , p_ud_ModulePathCompLen_Max  := #ud_ListHeaderPathCompLen_Max
                                , us_SDOMaxDataSize           := us_DataLength_Max
                                );

    //no response, error
    if ( sd_retval <> 0 ) then
      LogError("@ZZZZ (SafetyCDIAS_Base::ReadSDOConfig) Config Read Error: Error reading module path out of config data");
      return;
    end_if;

    // remember our own uncompressed path (first listheader path in the memory)
    if pListHeader^.p_us_Path & (GotOwnPath = FALSE) then
      GotOwnPath := TRUE;

      // remember the path
      _memcpy(ptr1:=#PathOfThisCPU[0], ptr2:=pListHeader^.p_us_Path, cntr:=(pListHeader^.p_us_Path$^UINT)^ + 2);
    end_if;

    //read length of download data in list-header (=LengthOverall) and save address
    //to calculate later the address of next list-header
    //address = last address + 4 byte (CRC)
    ud_ListLength_Address := ud_ListBaseAddress + 4;

    //send request and receive data
    sd_retval := SDOReadCfgRequ ( p_SDORequestBuffer  := p_SDORequestBuffer
                                , p_SDOResponseBuffer := p_SDOResponseBuffer
                                , ud_Address          := ud_ListLength_Address
                                , us_Length           := 4
                                );

    //no response
    if ( sd_retval <> 0 ) then
      LogError("@ZZZZ (SafetyCDIAS_Base::ReadSDOConfig) Config Read Error: Failed to read out the length of the download data within the configuration");
      return;
    end_if;

    //save length of list
    ud_ListLength := p_SDOResponseBuffer^.ud_Data;

    //read first opcode in interpreter list

    //                                                   v
    //address of LengthOverall + 4 bytes (LengthOverall, BlockType, ModuleID)
    ud_Address := ud_ListLength_Address + 4;

    // get BlockType
    //send request and receive data
    sd_retval := SDOReadCfgRequ ( p_SDORequestBuffer  := p_SDORequestBuffer
                                , p_SDOResponseBuffer := p_SDOResponseBuffer
                                , ud_Address          := ud_Address
                                , us_Length           := 4
                                );
    //no response, error
    if ( sd_retval <> 0 ) then
      LogError("@ZZZZ (SafetyCDIAS_Base::ReadSDOConfig) Config Read Error: Error getting the block type");
      return;
    end_if;

    ud_ActBlockType := p_SDOResponseBuffer^.ud_Data;

    case ud_ActBlockType of
//**********************************************************************************************************************************************************
      BLKTYPE_CFG_CPU,
      BLKTYPE_CFG_CPU_OPTIONAL , // if we don't need data from an external cpu
      BLKTYPE_CFG_MASTER_CPU:
        //add other CPUs to routing table

        // if there is a valid module path
        if pListHeader^.p_us_Path <> NIL then
          //add module to routing tabs
          sd_retval := AddModuleToRoutingTabs ( pModule       := pListHeader
                                              , pListHeader   := pListHeader
                                              , b_IsOptional  := (ud_ActBlockType = BLKTYPE_CFG_CPU_OPTIONAL)
                                              );

          if (sd_retval <> 0 ) then
            if ( ClassState <> _ModFromCfgNotFound ) then
              LogError("@ZZZZ (SafetyCDIAS_Base::ReadSDOConfig) Config Read Error: Failed to add cpu module to routing tabs");
              return;
            end_if;
          end_if;
        end_if;

//**********************************************************************************************************************************************************
      BLKTYPE_CFG_SLAVE_COMPR,
      BLKTYPE_CFG_SLAVE_COMPR_OPTIONAL: //Blocktyp der über die komprimierte Gesamtkonfiguration einer Slave-CPU gegeben wird
        //add other CPUs to routing table

        // if there is a valid module path
        if pListHeader^.p_us_Path <> NIL then
          //add module to routing tabs
          sd_retval := AddModuleToRoutingTabs ( pModule       := pListHeader
                                              , pListHeader   := pListHeader
                                              , b_IsOptional  := (ud_ActBlockType = BLKTYPE_CFG_SLAVE_COMPR_OPTIONAL)
                                              );

          if (sd_retval <> 0 ) then
            if ( ClassState <> _ModFromCfgNotFound ) then
              LogError("@ZZZZ (SafetyCDIAS_Base::ReadSDOConfig) Slave Config Read Error: Failed to add cpu module to routing tabs");
              return;
            end_if;
          end_if;

          // we skip the config till we get to the interface information of this slave (if it's the source of an interface frame we have to remember it)

          //address of LengthOverall + 3 * 4 bytes (LengthOverall, BlockType, ModuleID) => now the address points to FUB offset
          ud_Address := ud_ListLength_Address + 12;

          //skip FUB offset
          ud_Address += 4;

          // get no of FUB´s
          //send request and receive data
          sd_retval := SDOReadCfgRequ ( p_SDORequestBuffer  := p_SDORequestBuffer
                                      , p_SDOResponseBuffer := p_SDOResponseBuffer
                                      , ud_Address          := ud_Address
                                      , us_Length           := 4
                                      );
          //no response, error
          if ( sd_retval <> 0 ) then
            LogError("@ZZZZ (SafetyCDIAS_Base::ReadSDOConfig) Slave Config Read Error: Error getting the FUB number");
            return;
          end_if;

          ud_TmpCnt := p_SDOResponseBuffer^.ud_Data;

          // skip no of FUB´s and FUB´s
          ud_Address += (4 + (ud_TmpCnt * 4));

          // get length of path
          //send request and receive data
          sd_retval := SDOReadCfgRequ ( p_SDORequestBuffer  := p_SDORequestBuffer
                                      , p_SDOResponseBuffer := p_SDOResponseBuffer
                                      , ud_Address          := ud_Address
                                      , us_Length           := 4
                                      );
          //no response, error
          if ( sd_retval <> 0 ) then
            LogError("@ZZZZ (SafetyCDIAS_Base::ReadSDOConfig) Slave Config Read Error: Error getting the path length");
            return;
          end_if;

          ud_TmpCnt := p_SDOResponseBuffer^.ud_Data;

          // skip length of path and the path
          ud_Address += (4 + ud_TmpCnt);

          // get length of comp path
          //send request and receive data
          sd_retval := SDOReadCfgRequ ( p_SDORequestBuffer  := p_SDORequestBuffer
                                      , p_SDOResponseBuffer := p_SDOResponseBuffer
                                      , ud_Address          := ud_Address
                                      , us_Length           := 4
                                      );
          //no response, error
          if ( sd_retval <> 0 ) then
            LogError("@ZZZZ (SafetyCDIAS_Base::ReadSDOConfig) Slave Config Read Error: Error getting the comp path length");
            return;
          end_if;

          ud_TmpCnt := p_SDOResponseBuffer^.ud_Data;

          // skip length of comp path and the comp path
          ud_Address += (4 + ud_TmpCnt);

          // skip CRC and LengthOverall to get to the Blocktyp (Modul-Downloaddaten)
          ud_Address += 8;

          // get the block type
          //send request and receive data
          sd_retval := SDOReadCfgRequ ( p_SDORequestBuffer  := p_SDORequestBuffer
                                      , p_SDOResponseBuffer := p_SDOResponseBuffer
                                      , ud_Address          := ud_Address
                                      , us_Length           := 4
                                      );
          //no response, error
          if ( sd_retval <> 0 ) then
            LogError("@ZZZZ (SafetyCDIAS_Base::ReadSDOConfig) Slave Config Read Error: Error getting the block type of a slave config");
            return;
          end_if;

          ud_TmpCnt := p_SDOResponseBuffer^.ud_Data;

          // check if it's a new version of the configuration
          if (ud_TmpCnt = BLKTYPE_CFG_CONTAINER_V3)       |
             (ud_TmpCnt = BLKTYPE_CFG_CONTAINER_V3_SLAVE)     |
             (ud_TmpCnt = BLKTYPE_CFG_CONTAINER_V3_SLAVE_OPTIONAL) then

            // skip blocktype to get to the dynamic header length (how many data are attached to the header)
            ud_Address += 4;

            //send request and receive data
            sd_retval := SDOReadCfgRequ ( p_SDORequestBuffer  := p_SDORequestBuffer
                                        , p_SDOResponseBuffer := p_SDOResponseBuffer
                                        , ud_Address          := ud_Address
                                        , us_Length           := 4
                                        );

            //no response
            if ( sd_retval <> 0 ) then
              LogError("@ZZZZ (SafetyCDIAS_Base::ReadSDOConfig) Config Read Error: Error reading length of dynamic header data of a slave config");
              return;
            end_if;

            // plausibility check for data length
            if p_SDOResponseBuffer^.ud_Data > 1000 then
              sd_retval := -1;
              LogError("@ZZZZ (SafetyCDIAS_Base::ReadSDOConfig) Config Read Error: Invalid length of dynamic header data of a slave config");
              return;
            end_if;

            // the length info contains: size of length info + size of time info + size of additional data

            // skip the additional data to get to the path length
            ud_Address += p_SDOResponseBuffer^.ud_Data;
          else
            // old version => no dynamic header, so we skip only blocktype and time info
            ud_Address += 8;
          end_if;

          // get the path length
          //send request and receive data
          sd_retval := SDOReadCfgRequ ( p_SDORequestBuffer  := p_SDORequestBuffer
                                      , p_SDOResponseBuffer := p_SDOResponseBuffer
                                      , ud_Address          := ud_Address
                                      , us_Length           := 4
                                      );
          //no response, error
          if ( sd_retval <> 0 ) then
            LogError("@ZZZZ (SafetyCDIAS_Base::ReadSDOConfig) Slave Config Read Error: Error getting the path length");
            return;
          end_if;

          ud_TmpCnt := p_SDOResponseBuffer^.ud_Data;

          // skip length of path and the path
          ud_Address += (4 + ud_TmpCnt);

          // get length of comp path
          //send request and receive data
          sd_retval := SDOReadCfgRequ ( p_SDORequestBuffer  := p_SDORequestBuffer
                                      , p_SDOResponseBuffer := p_SDOResponseBuffer
                                      , ud_Address          := ud_Address
                                      , us_Length           := 4
                                      );
          //no response, error
          if ( sd_retval <> 0 ) then
            LogError("@ZZZZ (SafetyCDIAS_Base::ReadSDOConfig) Slave Config Read Error: Error getting the comp path length");
            return;
          end_if;

          ud_TmpCnt := p_SDOResponseBuffer^.ud_Data;

          // skip length of comp path and the comp path
          ud_Address += (4 + ud_TmpCnt);

          // skip CRC, LengthOverall, Blocktyp (Modul-Downloaddaten), ModuleID
          ud_Address += 16;

          // get the InterfaceCRC
          //send request and receive data
          sd_retval := SDOReadCfgRequ ( p_SDORequestBuffer  := p_SDORequestBuffer
                                      , p_SDOResponseBuffer := p_SDOResponseBuffer
                                      , ud_Address          := ud_Address
                                      , us_Length           := 4
                                      );
          //no response, error
          if ( sd_retval <> 0 ) then
            LogError("@ZZZZ (SafetyCDIAS_Base::ReadSDOConfig) Slave Config Read Error: Error getting the Inteface-CRC");
            return;
          end_if;

          TmpCRC := p_SDOResponseBuffer^.ud_Data;

          //add slave information to config
          AddSlaveToCfg ( pModule       := pListHeader
                        , b_IsOptional  := (ud_ActBlockType = BLKTYPE_CFG_SLAVE_COMPR_OPTIONAL)
                        , b_IsInterface := (TmpCRC <> 0)
                        , InterfaceCRC  := TmpCRC
                        );

        end_if;

//**********************************************************************************************************************************************************
      BLKTYPE_CFG_REV: // revision

        // check if the list is long enough for a String (more bytes than just the header)
        if ud_ListLength > 12 then

          //address of LengthOverall + 3 * 4 bytes (LengthOverall, BlockType, ModuleID) => now the address points to the revision string
          ud_Address := ud_ListLength_Address + 12;

          //read out the string (length = LengthOverall - length header)

          // get memory for the string
          if pPrjNameStr = NIL then
            PrjNameMemLen := ud_ListLength$USINT - 12;
            pPrjNameStr$^void := To_StdLib.Malloc(size := PrjNameMemLen + 1);
          else
            if PrjNameMemLen <> (ud_ListLength$USINT - 12) then
              PrjNameMemLen := ud_ListLength$USINT - 12;
              pPrjNameStr$^void := To_StdLib.ReAlloc(mptr:=pPrjNameStr, newsize:=PrjNameMemLen + 1);
            end_if;
          end_if;

          // check if we got a memory
          if pPrjNameStr then

            _memset(dest:=pPrjNameStr, usByte:=0, cntr:=PrjNameMemLen+1);

            ud_ActStrLen  := ud_TmpStrLen := PrjNameMemLen;
            ud_TmpAddress := ud_Address;

            IF p_BlockedTransferMemory = NIL THEN
              sd_retval   := -100;
              ClassState  := _MemAllocFailed;
              RETURN;
            END_IF;

            IF ud_BlockedTransferMemorySize < (ud_TmpStrLen + 1) THEN
              p_BlockedTransferMemory := To_StdLib.ReAlloc(mptr:=p_BlockedTransferMemory, newsize:=(ud_TmpStrLen + 1));
              IF p_BlockedTransferMemory = NIL THEN
                ud_BlockedTransferMemorySize  := 0;
                sd_retval                     := -100;
                ClassState                    := _MemAllocFailed;
                RETURN;
              ELSE
                ud_BlockedTransferMemorySize  := (ud_TmpStrLen + 1);
              END_IF;
            END_IF;

            To_StdLib.MemSet(dest:=p_BlockedTransferMemory, value:=0, size:=ud_BlockedTransferMemorySize);

            p_TmpBlockedData := p_BlockedTransferMemory;

            us_BlockedTransferLength := BlockedTransferLength(ud_Datalength:=ud_TmpStrLen, us_MaxBlocklength:=60);

            while us_BlockedTransferLength do

              // get name
              sd_retval := SDOReadCfgRequ ( p_SDORequestBuffer  := p_SDORequestBuffer
                                          , p_SDOResponseBuffer := p_SDOResponseBuffer
                                          , ud_Address          := ud_TmpAddress
                                          , us_Length           := us_BlockedTransferLength
                                          );
              //no response
              if ( sd_retval <> 0 ) then
                LogError("@ZZZZ (SafetyCDIAS_Base::ReadSDOConfig) Revision Read Error: Reading Revision failed");
                return;
              end_if;

              To_StdLib.MemCpy(dest   := p_TmpBlockedData,
                               source := #p_SDOResponseBuffer^.ud_Data,
                               size   := us_BlockedTransferLength);

              p_TmpBlockedData  += us_BlockedTransferLength;
              ud_TmpAddress     += us_BlockedTransferLength;
              ud_TmpStrLen      -= us_BlockedTransferLength;

              us_BlockedTransferLength := BlockedTransferLength(ud_Datalength:=ud_TmpStrLen, us_MaxBlocklength:=60);

            end_while;

            To_StdLib.MemCpy(dest   := pPrjNameStr,
                             source := p_BlockedTransferMemory,
                             size   := PrjNameMemLen+1);

            b_GotNewRevision  := TRUE;

            // string is formed by: project name {TAB} project revision   => search for the tab
            pPrjRevStr        := pPrjNameStr; // initialize pointer, because maybe there is no content in the projectname
            pChar             := pPrjNameStr;
            while pChar^ do
              // check for tab sign
              if pChar^ = 9 then
                // at the next character our revision starts
                pPrjRevStr    := pChar + sizeof(CHAR);

                // we change the tab to a string termination
                pChar^        := 0;

                // save the length of the name and the length of the project revision
                PrjNameStrLen := pChar$UDINT - pPrjNameStr$UDINT;
                PrjRevStrLen  := PrjNameMemLen - PrjNameStrLen - sizeof(CHAR);
                exit;
              end_if;

              pChar += sizeof(CHAR);
            end_while;

            ShowProjectRevision();
          end_if;
        end_if;

//**********************************************************************************************************************************************************
      BLKTYPE_CFG_INTERFACE,
      BLKTYPE_CFG_INTERFACE_OPTIONAL: // interface frame

        //address of LengthOverall + 3 * 4 bytes (LengthOverall, BlockType, Module ID) => points to interface CRC
        ud_Address := ud_ListLength_Address + 12;

//*****************************************************************************
//**   INTERFACE CRC                                                         **
//*****************************************************************************

        //send request and receive data
        sd_retval := SDOReadCfgRequ ( p_SDORequestBuffer  := p_SDORequestBuffer
                                    , p_SDOResponseBuffer := p_SDOResponseBuffer
                                    , ud_Address          := ud_Address
                                    , us_Length           := 4
                                    );

        //no response
        if ( sd_retval <> 0 ) then
          LogError("@ZZZZ (SafetyCDIAS_Base::ReadSDOConfig) Interface Config Read Error: Reading interface CRC of interface frame block failed");
          return;
        end_if;

        TempPdoConfig.InterfaceCRC := p_SDOResponseBuffer^.ud_Data;

        // skip interface crc
        ud_Address += 4;

//*****************************************************************************
//**   LENGTH OF TOPOLOGY PATH OF INTERFACE FRAME                            **
//*****************************************************************************

        //send request and receive data
        sd_retval := SDOReadCfgRequ ( p_SDORequestBuffer  := p_SDORequestBuffer
                                    , p_SDOResponseBuffer := p_SDOResponseBuffer
                                    , ud_Address          := ud_Address
                                    , us_Length           := 4
                                    );

        //no response
        if ( sd_retval <> 0 ) then
          LogError("@ZZZZ (SafetyCDIAS_Base::ReadSDOConfig) Interface Config Read Error: Reading length of topology path of interface frame block failed");
          return;
        end_if;

        // skip path length
        ud_Address += 4;

        us_BlockedTransferLength := p_SDOResponseBuffer^.ud_Data$USINT;

//*****************************************************************************
//**   TOPOLOGY PATH OF INTERFACE FRAME                                      **
//*****************************************************************************

        //send request and receive data
        sd_retval := SDOReadCfgRequ ( p_SDORequestBuffer  := p_SDORequestBuffer
                                    , p_SDOResponseBuffer := p_SDOResponseBuffer
                                    , ud_Address          := ud_Address
                                    , us_Length           := us_BlockedTransferLength
                                    );

        //no response
        if ( sd_retval <> 0 ) then
          LogError("@ZZZZ (SafetyCDIAS_Base::ReadSDOConfig) Interface Config Read Error: Reading topology path of interface frame block failed");
          return;
        end_if;

        // remember the destination path
        _memcpy(ptr1:=#TempPath[0], ptr2:=#p_SDOResponseBuffer^.ud_Data, cntr:=us_BlockedTransferLength);

        // skip path
        ud_Address += us_BlockedTransferLength;

//*****************************************************************************
//**   LENGTH OF COMPRESSED TOPOLOGY PATH OF INTERFACE FRAME                 **
//*****************************************************************************

        //send request and receive data
        sd_retval := SDOReadCfgRequ ( p_SDORequestBuffer  := p_SDORequestBuffer
                                    , p_SDOResponseBuffer := p_SDOResponseBuffer
                                    , ud_Address          := ud_Address
                                    , us_Length           := 4
                                    );

        //no response
        if ( sd_retval <> 0 ) then
          LogError("@ZZZZ (SafetyCDIAS_Base::ReadSDOConfig) Interface Config Read Error: Reading length of compressed topology path of interface frame block failed");
          return;
        end_if;

        // skip path length
        ud_Address += 4;

        us_BlockedTransferLength := p_SDOResponseBuffer^.ud_Data$USINT;

//*****************************************************************************
//**   COMPRESSED TOPOLOGY PATH OF INTERFACE FRAME                           **
//*****************************************************************************

        //send request and receive data
        sd_retval := SDOReadCfgRequ ( p_SDORequestBuffer  := p_SDORequestBuffer
                                    , p_SDOResponseBuffer := p_SDOResponseBuffer
                                    , ud_Address          := ud_Address
                                    , us_Length           := us_BlockedTransferLength
                                    );

        //no response
        if ( sd_retval <> 0 ) then
          LogError("@ZZZZ (SafetyCDIAS_Base::ReadSDOConfig) Interface Config Read Error: Reading compressed topology path of interface frame block failed");
          return;
        end_if;

        // skip path and maximum cycle time
        ud_Address += us_BlockedTransferLength + 4;

  // here starts the data area (before we read only the list header

//*****************************************************************************
//**   INTERFACE CRC                                                         **
//*****************************************************************************

        //send request and receive data
        sd_retval := SDOReadCfgRequ ( p_SDORequestBuffer  := p_SDORequestBuffer
                                    , p_SDOResponseBuffer := p_SDOResponseBuffer
                                    , ud_Address          := ud_Address
                                    , us_Length           := 4
                                    );

        //no response
        if ( sd_retval <> 0 ) then
          LogError("@ZZZZ (SafetyCDIAS_Base::ReadSDOConfig) Interface Config Read Error: Reading CRC of interface frame block failed");
          return;
        end_if;

        TempPdoConfig.InterfaceCRC := p_SDOResponseBuffer^.ud_Data;

        // skip interface CRC
        ud_Address += 4;

//*****************************************************************************
//**   NUMBER OF BOOL INTERFACE VARIABLES IN THE PDO                         **
//*****************************************************************************

        //send request and receive data
        sd_retval := SDOReadCfgRequ ( p_SDORequestBuffer  := p_SDORequestBuffer
                                    , p_SDOResponseBuffer := p_SDOResponseBuffer
                                    , ud_Address          := ud_Address
                                    , us_Length           := 4
                                    );

        //no response
        if ( sd_retval <> 0 ) then
          LogError("@ZZZZ (SafetyCDIAS_Base::ReadSDOConfig) Interface Config Read Error: Reading number of bool variables in the interface frame failed");
          return;
        end_if;

        BoolOuts := p_SDOResponseBuffer^.ud_Data;

        // skip bool variables
        ud_Address += 4;

//*****************************************************************************
//**   NUMBER OF DINT INTERFACE VARIABLES IN THE PDO                         **
//*****************************************************************************

        //send request and receive data
        sd_retval := SDOReadCfgRequ ( p_SDORequestBuffer  := p_SDORequestBuffer
                                    , p_SDOResponseBuffer := p_SDOResponseBuffer
                                    , ud_Address          := ud_Address
                                    , us_Length           := 4
                                    );

        //no response
        if ( sd_retval <> 0 ) then
          LogError("@ZZZZ (SafetyCDIAS_Base::ReadSDOConfig) Interface Config Read Error: Reading number of dint variables in the interface frame failed");
          return;
        end_if;

        // skip bool variables
        ud_Address += 4;

        DintOuts := p_SDOResponseBuffer^.ud_Data;

        // if there are interface variables
        if BoolOuts | DintOuts then
          // calculate the length of the interface frame
          TempPdoConfig.PdoLen              := CalcPDOLength(BoolOuts, DintOuts);

          // this is the source of the interface frame
          TempPdoConfig.SourcePathLen       := TempPath[0]$UINT + 2;
          TempPdoConfig.pSourcePath         := #TempPath[0];

          // and the destination
          TempPdoConfig.DestPathLen         := PathOfThisCPU[0]$UINT + 2;
          TempPdoConfig.pDestPath           := #PathOfThisCPU[0];

          TempPdoConfig.Info                := 0;
          TempPdoConfig.Info.IsInterfacePDO := TRUE;
          TempPdoConfig.Info.IsOptional     := (ud_ActBlockType = BLKTYPE_CFG_INTERFACE_OPTIONAL);

          // add the interface PDO to the list
          AddPdoToCfg(TempPdoConfig);
        else
          LogError("@ZZZZ (SafetyCDIAS_Base::ReadSDOConfig) Interface Config Read Error: No interface variables found in interface blocktype");
          return;
        end_if;

//**********************************************************************************************************************************************************
      BLKTYPE_CFG_MODULE,
      BLKTYPE_CFG_MODULE_V2,
      BLKTYPE_CFG_MODULE_OPTIONAL,
      BLKTYPE_CFG_CONTAINER_SLAVE,
      BLKTYPE_CFG_CONTAINER_SLAVE_OPTIONAL,
      BLKTYPE_CFG_MODULE_V3,
      BLKTYPE_CFG_MODULE_V3_OPTIONAL,
      BLKTYPE_CFG_CONTAINER_V3_SLAVE,
      BLKTYPE_CFG_CONTAINER_V3_SLAVE_OPTIONAL:      // module configurations
        TempModuleConfig.Info               := 0;
        TempModuleConfig.DestCRCNo          := 0;
        TempModuleConfig.pDestCRCs          := NIL;
        if ud_ActBlockType = BLKTYPE_CFG_MODULE_OPTIONAL then
          TempModuleConfig.Info.IsOptional  := TRUE;
        else
          TempModuleConfig.Info.IsOptional  := FALSE;
        end_if;

        b_CfgTypeV2 := (ud_ActBlockType <> BLKTYPE_CFG_MODULE);

        // check if it's a V3 config, because the structure of the IO List is different
        if (ud_ActBlockType = BLKTYPE_CFG_MODULE_V3) |
           (ud_ActBlockType = BLKTYPE_CFG_MODULE_V3_OPTIONAL) |
           (ud_ActBlockType = BLKTYPE_CFG_CONTAINER_V3_SLAVE) |
           (ud_ActBlockType = BLKTYPE_CFG_CONTAINER_V3_SLAVE_OPTIONAL) then
          b_CfgTypeV3 := TRUE;
        else
          b_CfgTypeV3 := FALSE;
        end_if;

        // if it's our own path, remember the type of module configuration
        if (PathOfThisCPU[0]$UINT = (pListHeader^.p_us_Path$^UINT)^) & (To_StdLib.MemCmp(#PathOfThisCPU[0], pListHeader^.p_us_Path, PathOfThisCPU[0]$UINT + 2) = 0) then
          // if config is already "old" dont change to "new". (can be set by block BLKTYPE_OLD_MODE_FLAG)
          if NewConfigType <> ConfigState_Old then
            NewConfigType := (b_CfgTypeV2$USINT + 1)$t_ConfigStateType;
          end_if;
        end_if;

        BoolOuts := 0;
        DintOuts := 0;

        // Remember the path (uncompressed and compressed)
        TempModuleConfig.PathLen      := pListHeader^.p_us_Path^$UINT + 2;
        TempModuleConfig.pPath        := pListHeader^.p_us_Path;

        TempModuleConfig.CompPathLen  := pListHeader^.ui_PathCompLen;
        TempModuleConfig.pCompPath    := pListHeader^.p_us_PathComp;

//*****************************************************************************
//**   LIST HEADER                                                           **
//*****************************************************************************

        //address of LengthOverall + 3 * 4 bytes (LengthOverall, BlockType, ModuleID)
        ud_Address := ud_ListLength_Address + 12;

        // only available at new modules
        if b_CfgTypeV2 then

//*****************************************************************************
//**   INTERFACE CRC                                                         **
//*****************************************************************************

          //send request and receive data
          sd_retval := SDOReadCfgRequ ( p_SDORequestBuffer  := p_SDORequestBuffer
                                      , p_SDOResponseBuffer := p_SDOResponseBuffer
                                      , ud_Address          := ud_Address
                                      , us_Length           := 4
                                      );

          //no response
          if ( sd_retval <> 0 ) then
            LogError("@ZZZZ (SafetyCDIAS_Base::ReadSDOConfig) Config Read Error: Reading interface CRC of interface frame block failed");
            return;
          end_if;

          TempPdoConfig.InterfaceCRC := p_SDOResponseBuffer^.ud_Data;

          // skip interface crc
          ud_Address += 4;

//*****************************************************************************
//**   LENGTH OF TOPOLOGY PATH OF INTERFACE FRAME                            **
//*****************************************************************************

          //send request and receive data
          sd_retval := SDOReadCfgRequ ( p_SDORequestBuffer  := p_SDORequestBuffer
                                      , p_SDOResponseBuffer := p_SDOResponseBuffer
                                      , ud_Address          := ud_Address
                                      , us_Length           := 4
                                      );

          //no response
          if ( sd_retval <> 0 ) then
            LogError("@ZZZZ (SafetyCDIAS_Base::ReadSDOConfig) Config Read Error: Reading length of topology path of interface frame block failed");
            return;
          end_if;

          // skip path length
          ud_Address += 4;

          us_BlockedTransferLength := p_SDOResponseBuffer^.ud_Data$USINT;

//*****************************************************************************
//**   TOPOLOGY PATH OF INTERFACE FRAME                                      **
//*****************************************************************************

          //send request and receive data
          sd_retval := SDOReadCfgRequ ( p_SDORequestBuffer  := p_SDORequestBuffer
                                      , p_SDOResponseBuffer := p_SDOResponseBuffer
                                      , ud_Address          := ud_Address
                                      , us_Length           := us_BlockedTransferLength
                                      );

          //no response
          if ( sd_retval <> 0 ) then
            LogError("@ZZZZ (SafetyCDIAS_Base::ReadSDOConfig) Config Read Error: Reading topology path of interface frame block failed");
            return;
          end_if;

          // remember the destination path
          _memcpy(ptr1:=#TempPath[0], ptr2:=#p_SDOResponseBuffer^.ud_Data, cntr:=us_BlockedTransferLength);

          // skip path
          ud_Address += us_BlockedTransferLength;

//*****************************************************************************
//**   LENGTH OF COMPRESSED TOPOLOGY PATH OF INTERFACE FRAME                 **
//*****************************************************************************

          //send request and receive data
          sd_retval := SDOReadCfgRequ ( p_SDORequestBuffer  := p_SDORequestBuffer
                                      , p_SDOResponseBuffer := p_SDOResponseBuffer
                                      , ud_Address          := ud_Address
                                      , us_Length           := 4
                                      );

          //no response
          if ( sd_retval <> 0 ) then
            LogError("@ZZZZ (SafetyCDIAS_Base::ReadSDOConfig) Config Read Error: Reading length of compressed topology path of interface frame block failed");
            return;
          end_if;

          // skip path length
          ud_Address += 4;

          us_BlockedTransferLength := p_SDOResponseBuffer^.ud_Data$USINT;

//*****************************************************************************
//**   COMPRESSED TOPOLOGY PATH OF INTERFACE FRAME                           **
//*****************************************************************************

          //send request and receive data
          sd_retval := SDOReadCfgRequ ( p_SDORequestBuffer  := p_SDORequestBuffer
                                      , p_SDOResponseBuffer := p_SDOResponseBuffer
                                      , ud_Address          := ud_Address
                                      , us_Length           := us_BlockedTransferLength
                                      );

          //no response
          if ( sd_retval <> 0 ) then
            LogError("@ZZZZ (SafetyCDIAS_Base::ReadSDOConfig) Config Read Error: Reading compressed topology path of interface frame block failed");
            return;
          end_if;

          ud_Address += us_BlockedTransferLength;

          // skip max. cycle time
          ud_Address += 4;
        end_if;

        // on first 4 bytes is fix the system time
        ud_ActAddress := 4;

        // address in memory for unsafe BDINT variables
        ud_UnsafeBDINT_Offset := 0;

//*****************************************************************************
//**   INTERPRETER CODE                                                      **
//*****************************************************************************

        //read til end-command is reached
        while ( 1 ) do

          //send request and receive data
          sd_retval := SDOReadCfgRequ ( p_SDORequestBuffer  := p_SDORequestBuffer
                                      , p_SDOResponseBuffer := p_SDOResponseBuffer
                                      , ud_Address          := ud_Address
                                      , us_Length           := 4
                                      );
          //no response, error
          if ( sd_retval <> 0 ) then
            LogError("@ZZZZ (SafetyCDIAS_Base::ReadSDOConfig) Config Read Error: Reading next command failed");
            return;
          end_if;

          //end-command found
          if ( p_SDOResponseBuffer^.ud_Data = SDO_CONFIG_END_CMD ) then
            exit;
          end_if;

          //read next opcode
          //length of one command = 4 x 4 bytes
          ud_Address += 16;

          //if there is no end-command found, the returncode of response will be <> OK, when the end of config data is missed
          //In this case the loop ends with returncode <> 0.
        end_while;

        //list of I/Os starts at last address + 16 (length of end command = 4x4 bytes)
        ud_Address += 16;

//*****************************************************************************
//**   LOCAL BOOL INPUTS                                                     **
//*****************************************************************************

        //read number of local bool inputs

        //send request and receive data
        sd_retval := SDOReadCfgRequ ( p_SDORequestBuffer  := p_SDORequestBuffer
                                    , p_SDOResponseBuffer := p_SDOResponseBuffer
                                    , ud_Address          := ud_Address
                                    , us_Length           := 4
                                    );

        //no response
        if ( sd_retval <> 0 ) then
          LogError("@ZZZZ (SafetyCDIAS_Base::ReadSDOConfig) Config Read Error: Reading number of local inputs failed");
          return;
        end_if;

        // remember the number
        BoolOuts += p_SDOResponseBuffer^.ud_Data;

        // get offset in application memory
        ud_ActAddress += p_SDOResponseBuffer^.ud_Data * 4;

        //++pr
        ud_skipLength := 4; // Anzahl Einträge
        // only available at new modules
        if b_CfgTypeV2 then
          ud_skipLength += 12 * p_SDOResponseBuffer^.ud_Data; // QSE, Filtertime, Modulkennung(SDIAS)
        else
          ud_skipLength += 8 * p_SDOResponseBuffer^.ud_Data; // QSE, Filtertime
        end_if;

//*****************************************************************************
//**   LOCAL BOOL OUTPUTS AS INPUTS                                          **
//*****************************************************************************

        // get number of safe outputs as inputs

        //send request and receive data
        sd_retval := SDOReadCfgRequ ( p_SDORequestBuffer  := p_SDORequestBuffer
                                    , p_SDOResponseBuffer := p_SDOResponseBuffer
                                    , ud_Address          := p_SDORequestBuffer^.ud_Address + ud_skipLength // ++pr
                                    , us_Length           := 4
                                    );

        //no response
        if ( sd_retval <> 0 ) then
          LogError("@ZZZZ (SafetyCDIAS_Base::ReadSDOConfig) Config Read Error: Reading number of safe outputs as inputs failed");
          return;
        end_if;

        // remember the number
        BoolOuts += p_SDOResponseBuffer^.ud_Data;

        // get offset in application memory
        ud_ActAddress += p_SDOResponseBuffer^.ud_Data * 4;

//*****************************************************************************
//**   SAFE BOOL OUTPUT VARIABLES                                            **
//*****************************************************************************

        // get number of safe bool output vars

        //send request and receive data
        sd_retval := SDOReadCfgRequ ( p_SDORequestBuffer  := p_SDORequestBuffer
                                    , p_SDOResponseBuffer := p_SDOResponseBuffer
                                    , ud_Address          := p_SDORequestBuffer^.ud_Address + 4
                                    , us_Length           := 4
                                    );

        //no response
        if ( sd_retval <> 0 ) then
          LogError("@ZZZZ (SafetyCDIAS_Base::ReadSDOConfig) Config Read Error: Reading number of safe bool output vars failed");
          return;
        end_if;

        // remember the number
        BoolOuts += p_SDOResponseBuffer^.ud_Data;

        // get offset in application memory
        ud_ActAddress += p_SDOResponseBuffer^.ud_Data * 4;

        // the new container has some additional content here
        if b_CfgTypeV3 then

//*****************************************************************************
//**   LOCAL DINT INPUTS                                                     **
//*****************************************************************************

          //read number of local dint inputs

          //send request and receive data
          sd_retval := SDOReadCfgRequ ( p_SDORequestBuffer  := p_SDORequestBuffer
                                      , p_SDOResponseBuffer := p_SDOResponseBuffer
                                      , ud_Address          := p_SDORequestBuffer^.ud_Address + 4
                                      , us_Length           := 4
                                      );

          //no response
          if ( sd_retval <> 0 ) then
            LogError("@ZZZZ (SafetyCDIAS_Base::ReadSDOConfig) Config Read Error: Reading number of local DINT inputs failed");
            return;
          end_if;

          // remember the number
          DintOuts += p_SDOResponseBuffer^.ud_Data;

          // get offset in application memory
          ud_ActAddress += p_SDOResponseBuffer^.ud_Data * 4;

//*****************************************************************************
//**   LOCAL DINT OUTPUTS AS INPUTS                                          **
//*****************************************************************************

          // get number of safe dint outputs as inputs

          //send request and receive data
          sd_retval := SDOReadCfgRequ ( p_SDORequestBuffer  := p_SDORequestBuffer
                                      , p_SDOResponseBuffer := p_SDOResponseBuffer
                                      , ud_Address          := p_SDORequestBuffer^.ud_Address + 4 + 12 * p_SDOResponseBuffer^.ud_Data
                                      , us_Length           := 4
                                      );

          //no response
          if ( sd_retval <> 0 ) then
            LogError("@ZZZZ (SafetyCDIAS_Base::ReadSDOConfig) Config Read Error: Reading number of safe DINT outputs as inputs failed");
            return;
          end_if;

          // remember the number
          DintOuts += p_SDOResponseBuffer^.ud_Data;

          // get offset in application memory
          ud_ActAddress += p_SDOResponseBuffer^.ud_Data * 4;

        end_if;

//*****************************************************************************
//**   SAFE DINT OUTPUT VARIABLES                                            **
//*****************************************************************************

        // get number of safe dint output vars

        //send request and receive data
        sd_retval := SDOReadCfgRequ ( p_SDORequestBuffer  := p_SDORequestBuffer
                                    , p_SDOResponseBuffer := p_SDOResponseBuffer
                                    , ud_Address          := p_SDORequestBuffer^.ud_Address + 4
                                    , us_Length           := 4
                                    );

        //no response
        if ( sd_retval <> 0 ) then
          LogError("@ZZZZ (SafetyCDIAS_Base::ReadSDOConfig) Config Read Error: Reading number of safe dint output vars failed");
          return;
        end_if;

        // only when there is a manager
        if pSafetyManagerThis then
          // remember the number
          DintOuts += p_SDOResponseBuffer^.ud_Data;

          // now we're ready to determine the PDO size of this module
          TempModuleConfig.PdoOutLen := CalcPDOLength(BoolOuts, DintOuts);

          // if it's our own path, remember the PDO length
          if (PathOfThisCPU[0]$UINT = (pListHeader^.p_us_Path$^UINT)^) & (To_StdLib.MemCmp(#PathOfThisCPU[0], pListHeader^.p_us_Path, PathOfThisCPU[0]$UINT + 2) = 0) then
            MyPDOSize := TempModuleConfig.PdoOutLen;
          end_if;
        end_if;

        // get offset in application memory
        ud_ActAddress += p_SDOResponseBuffer^.ud_Data * 4;

        // special unsafe variables (not supported by old modules)
        if b_CfgTypeV2 then

//*****************************************************************************
//**   FAST UNSAFE OUTPUT VARIABLES                                          **
//*****************************************************************************

          // get number of fast unsafe output vars (should be 8 or 0)

          //send request and receive data
          sd_retval := SDOReadCfgRequ ( p_SDORequestBuffer  := p_SDORequestBuffer
                                      , p_SDOResponseBuffer := p_SDOResponseBuffer
                                      , ud_Address          := p_SDORequestBuffer^.ud_Address + 4
                                      , us_Length           := 4
                                      );

          //no response
          if ( sd_retval <> 0 ) then
            LogError("@ZZZZ (SafetyCDIAS_Base::ReadSDOConfig) Config Read Error: Reading number of fast unsafe output vars failed");
            return;
          end_if;

          // get offset in application memory
          ud_ActAddress += p_SDOResponseBuffer^.ud_Data * 4;
